(* Logix 5000 project; controller lab4BnB 5069-L306ERM rev 38.11; software revision 38.02 *)

TASK MainTask (periodic, rate 1 ms, priority 10, watchdog 1 ms) : MainProgram

MODULES
   Local : 5069-L306ERM (5069 0, rev 38.11)
       : vendor 1 type 115 code 320 (5069 4, rev 2.13, StandardDataDriven RPI 1 ms)
       : 5069-IF8 (5069 3, rev 3.11, StandardDataDriven RPI 1 ms)
       : 5069-IB16 (5069 1, rev 2.16, StandardDataDriven RPI 5 ms)
       : 5069-OB16 (5069 2, rev 3.13, StandardDataDriven RPI 5 ms)
END_MODULES

VAR_GLOBAL   (* controller tags *)
   BalanceMax : REAL := 2.8;
   BalanceMin : REAL := -1.92;
   DesiredMotorAngleDeg : DINT := 45;
   Kd : REAL := 0.8;
   Ki : REAL := 0.5;
   Kp : REAL := 0.5;
   MotorAngleDeg : DINT := 45;
   MotorInInt : ALIAS FOR Local:4:O.Ch00.Data;
   MotorVoltageInt : ALIAS FOR Local:3:I.Ch00.Data;
   MyError : DINT;
   PostFilter : DINT;
   PreFilter : DINT;
END_VAR

PROGRAM MainProgram   (* main routine main *)
VAR
   DERV_01 : DERIVATIVE := (Gain := 0.8, RTSTime := 1, DeltaT := 0.001);
   INTG_02 : INTEGRATOR := (IGain := 0.5, HighLimit := 4.0, LowLimit := -4.0, RTSTime := 1, Out := -0.06536653, DeltaT := 0.001);
   LPF_01 : FILTER_LOW_PASS := (WLag := 0.5, Order := 1, RTSTime := 1, DeltaT := 0.001);
   MUL_01 : FBD_MATH := (SourceA := 0.5);
   SCL_01 : SCALE := (In := 1.6302257, InRawMax := 2.8, InRawMin := -1.92, InEUMax := 90.0, InEUMin := -90.0, Limiting := 1, Out := 45.38997);
   SCL_02 : SCALE := (In := -0.06536653, InRawMax := 90.0, InRawMin := -90.0, InEUMax := -10.0, InEUMin := 10.0, Limiting := 1, Out := 0.0072631836);
   SSUM_01 : SELECTED_SUMMER := (Gain1 := 1.0, Select1 := 1, Gain2 := 1.0, Select2 := 1, In3 := -0.06536653, Gain3 := 1.0, Select3 := 1, Gain4 := 1.0, Gain5 := 1.0, Gain6 := 1.0, Gain7 := 1.0, Gain8 := 1.0, Out := -0.06536653);
   SUB_01 : FBD_MATH := (SourceA := 45.0, SourceB := 45.0);
END_VAR

ROUTINE main   (* function block diagram *)
   SHEET 1
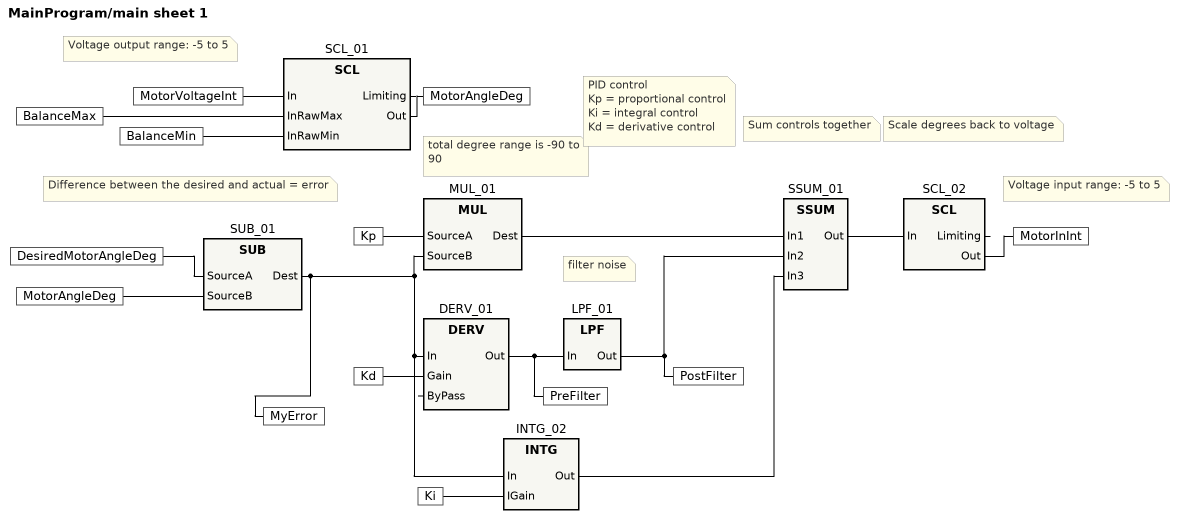
   // Difference between the desired and actual = error
   // Voltage output range: -5 to 5
   // total degree range is -90 to
   // 90
   // filter noise
   // PID control
   // Kp = proportional control
   // Ki = integral control
   // Kd = derivative control
   // Sum controls together
   // Scale degrees back to voltage
   // Voltage input range: -5 to 5
   SUB_01 : SUB(SourceA := DesiredMotorAngleDeg, SourceB := MotorAngleDeg);
   MyError := SUB_01.Dest;
   SCL_01 : SCL(In := MotorVoltageInt, InRawMax := BalanceMax, InRawMin := BalanceMin);   // unwired pins: Limiting
   MotorAngleDeg := SCL_01.Out;
   MUL_01 : MUL(SourceA := Kp, SourceB := SUB_01.Dest);
   DERV_01 : DERV(In := SUB_01.Dest, Gain := Kd);   // unwired pins: ByPass
   INTG_02 : INTG(In := SUB_01.Dest, IGain := Ki);
   PreFilter := DERV_01.Out;
   LPF_01 : LPF(In := DERV_01.Out);
   PostFilter := LPF_01.Out;
   SSUM_01 : SSUM(In1 := MUL_01.Dest, In2 := LPF_01.Out, In3 := INTG_02.Out);
   SCL_02 : SCL(In := SSUM_01.Out);   // unwired pins: Limiting
   MotorInInt := SCL_02.Out;
END_ROUTINE
END_PROGRAM
